FUNCTION_BLOCK FB_SatelliteController IMPLEMENTS I_FeedLoad, I_JsonSource
VAR_INPUT
    stCfg : ST_BoxConfig;  // this box's row of GVL_Config.aBoxes
END_VAR
VAR_OUTPUT
    bValid      : BOOL;   // the values below can be used
    bMeasured   : BOOL;   // TRUE: from the supply. FALSE: estimated from the feed
    fDcAmps     : LREAL;  // A DC, filtered
    fDcVolts    : LREAL;  // V DC
    fAcPowerW   : LREAL;  // W on the AC side, at the box
    fCableLossW : LREAL;  // W lost in the box's own AC cable, on top of fAcPowerW
END_VAR
VAR
    fbSupply  : FB_EcPowerSupply;
    fEff      : LREAL := 0.95;
    fCycleS   : LREAL;
    fRawLossW : LREAL;  // cable loss from this cycle's unfiltered current
END_VAR

fEff    := LIMIT(0.5, stCfg.fPsuEfficiency, 1.0);
fCycleS := F_CycleTimeS();

IF stCfg.bHasEcPowerSupply THEN
    bMeasured := TRUE;
    fbSupply(bSimulate := GVL_Config.bSimulateSupplies);

    IF fbSupply.bOnline THEN
        fDcVolts  := fbSupply.fOutputVolts;
        // The loss goes with the square of the current, so it is taken from the raw current every cycle and
        // filtered afterwards. Filtering the current first would read low whenever the load moves.
        fRawLossW := F_CableLossW(fPowerW := fDcVolts * fbSupply.fOutputAmps / fEff,
                                  fLengthFt := stCfg.fWireLengthFt, nAwg := stCfg.nWireAwg);
        IF bValid THEN
            fDcAmps     := F_LowPass(fState := fDcAmps,     fInput := fbSupply.fOutputAmps, fTimeS := GVL_Config.fFilterTimeS, fCycleS := fCycleS);
            fCableLossW := F_LowPass(fState := fCableLossW, fInput := fRawLossW,            fTimeS := GVL_Config.fFilterTimeS, fCycleS := fCycleS);
        ELSE
            fDcAmps     := fbSupply.fOutputAmps;  // first valid sample: no filter run-in
            fCableLossW := fRawLossW;
        END_IF
        fAcPowerW := fDcVolts * fDcAmps / fEff;
        bValid    := TRUE;
    ELSE
        // Off the bus: counted as 0 W and reported as not valid.
        fDcAmps     := 0.0;
        fDcVolts    := 0.0;
        fAcPowerW   := 0.0;
        fCableLossW := 0.0;
        bValid      := FALSE;
    END_IF
ELSE
    // No supply: SetShare() writes the outputs when the feed has done its split.
    bMeasured := FALSE;
END_IF

METHOD GetDemand : ST_LoadDemand
VAR
    stDemand : ST_LoadDemand;
END_VAR
// What the feed sees at the branch point: the box's draw plus the loss in the box's cable.
stDemand.fCableFactor := F_CableFactor(fLengthFt := stCfg.fWireLengthFt, nAwg := stCfg.nWireAwg);
IF stCfg.bHasEcPowerSupply THEN
    stDemand.eKind       := E_LoadKind.Measured;
    stDemand.fAcPowerW   := fAcPowerW + fCableLossW;
    stDemand.fCableLossW := fCableLossW;
    stDemand.fWeight     := 0.0;
    stDemand.bValid      := bValid;
ELSE
    stDemand.eKind       := E_LoadKind.Estimated;
    stDemand.fAcPowerW   := 0.0;
    stDemand.fCableLossW := fCableLossW;  // from the share, once SetShare() has run this cycle
    stDemand.fWeight     := UDINT_TO_LREAL(stCfg.nPixelCount);
    stDemand.bValid      := TRUE;
END_IF
GetDemand := stDemand;
END_METHOD

METHOD SetShare
VAR_INPUT
    fShareW     : LREAL;  // W on the AC side
    bShareValid : BOOL;   // FALSE: the feed has no valid measurement
END_VAR
IF NOT stCfg.bHasEcPowerSupply THEN
    // The share includes the loss in the box's own cable. What arrives at the box is less.
    fAcPowerW   := F_PowerAfterCable(fShareW := fShareW, fLengthFt := stCfg.fWireLengthFt, nAwg := stCfg.nWireAwg);
    fCableLossW := MAX(0.0, fShareW) - fAcPowerW;
    fDcVolts    := stCfg.fNominalDcVolts;
    IF stCfg.fNominalDcVolts > 1.0 THEN
        fDcAmps := fAcPowerW * fEff / stCfg.fNominalDcVolts;
    ELSE
        fDcAmps := 0.0;
    END_IF
    bValid := bShareValid;
END_IF
END_METHOD

METHOD WriteJson
VAR_INPUT
    eSection : E_JsonSection;
END_VAR
VAR_IN_OUT
    fbJson : FB_JsonSaxWriter;
END_VAR
VAR
    sFeed : STRING(20);
END_VAR
IF eSection <> E_JsonSection.Box THEN
    RETURN;
END_IF

sFeed := F_FeedIdString(nFeedId := stCfg.nFeedId);

fbJson.AddKey('id');
fbJson.AddString(stCfg.sId);
fbJson.AddKey('name');
fbJson.AddString(stCfg.sControllerName);
fbJson.AddKey('feed');
fbJson.AddString(sFeed);
F_JsonInt(sKey := 'pixels', nValue := UDINT_TO_DINT(MIN(stCfg.nPixelCount, 2147483647)), fbJson := fbJson);
F_JsonNum(sKey := 'maxDcAmps', fValue := stCfg.fMaxDcCurrent, bValid := TRUE, nDecimals := 1, fbJson := fbJson);
fbJson.AddKey('src');
IF stCfg.bHasEcPowerSupply THEN
    fbJson.AddString('psu');
ELSE
    fbJson.AddString('est');
END_IF
fbJson.AddKey('ok');
fbJson.AddBool(bValid);
F_JsonNum(sKey := 'dcAmps', fValue := fDcAmps, bValid := bValid, nDecimals := 2, fbJson := fbJson);
F_JsonNum(sKey := 'dcVolts', fValue := fDcVolts, bValid := bValid AND stCfg.bHasEcPowerSupply, nDecimals := 1, fbJson := fbJson);
F_JsonNum(sKey := 'acW', fValue := fAcPowerW, bValid := bValid, nDecimals := 1, fbJson := fbJson);
F_JsonNum(sKey := 'cableLossW', fValue := fCableLossW, bValid := bValid, nDecimals := 1, fbJson := fbJson);

fbJson.AddKey('psu');
IF stCfg.bHasEcPowerSupply THEN
    fbJson.StartObject();
    fbJson.AddKey('dcOk');
    fbJson.AddBool(fbSupply.bDcOk);
    fbJson.AddKey('warn');
    fbJson.AddBool(fbSupply.bWarning);
    fbJson.AddKey('err');
    fbJson.AddBool(fbSupply.bError);
    F_JsonNumSigned(sKey := 'tempC', fValue := fbSupply.fTempC, bValid := fbSupply.bTempValid, nDecimals := 0, fbJson := fbJson);
    F_JsonNum(sKey := 'inVolts', fValue := fbSupply.fInputVolts, bValid := fbSupply.bInputVoltsValid, nDecimals := 0, fbJson := fbJson);
    fbJson.EndObject();
ELSE
    fbJson.AddNull();
END_IF
END_METHOD

END_FUNCTION_BLOCK

(* stored: Version 1.1.0.1
   POU FB_SatelliteController: Id {fd4bea5b-c411-438a-8000-f3f90d5fc734}, SpecialFunc None
   Method GetDemand: Id {f5bd97ef-6b3a-4a18-9fc2-a3a18bdf500d}
   Method SetShare: Id {19e24c6f-0ed2-426d-bffb-736a7c11d6c1}
   Method WriteJson: Id {b943426d-e14b-4302-a995-308542171dec} *)
